screen "Rack 2" 640x480
   Button "Button_1" at 0,0 size 90x66; TextOff 'Rack 1'
      on Click: ActivateScreen("Rack 1", 0)
   Button "Button_2" at 130,0 size 90x66; TextOff 'Rack 2'
      on Click: ActivateScreen("Rack 2", 0)
   DateTimeField "Date/time field_1" at 444,15 size 177x31
   TextField "Text field_46" at 350,88 size 74x28; Text 'Rack 2'
   ScreenModuleView "RackSlot_1" at 562,360 size 44x36; Guid_{11997190-21654} '0'; ScreenModuleType ""
      on Guid_{11997190-21491}: function_efd93a16("RackSlotData", 0, 0, -1, -1, 1)
      Guid_{11997190-21133} <- "WarehouseData_Rack1{1}"
   ScreenModuleView "RackSlot_2" at 512,360 size 44x36; Guid_{11997190-21654} '0'; ScreenModuleType ""
      on Guid_{11997190-21491}: function_efd93a16("RackSlotData", 0, 0, -1, -1, 1)
      Guid_{11997190-21133} <- "WarehouseData_Rack1{1}"
   ScreenModuleView "RackSlot_3" at 562,360 size 44x36; Guid_{11997190-21654} '1'; Guid_{11997190-23841} '1'; ScreenModuleType ""
      on Guid_{11997190-21491}: SetTag("SelectedRack", 2); SetTag("SelectedSlot", 1); function_efd93a16("RackSlotData", 220, 150, -1, -1, 1)
      Guid_{11997190-21133} <- "WarehouseData_Rack2{1}"
   ScreenModuleView "RackSlot_4" at 512,360 size 44x36; Guid_{11997190-21654} '2'; Guid_{11997190-23841} '2'; ScreenModuleType ""
      on Guid_{11997190-21491}: SetTag("SelectedRack", 2); SetTag("SelectedSlot", 2); function_efd93a16("RackSlotData", 220, 150, -1, -1, 1)
      Guid_{11997190-21133} <- "WarehouseData_Rack2{2}"
   ScreenModuleView "RackSlot_5" at 462,360 size 44x36; Guid_{11997190-21654} '3'; Guid_{11997190-23841} '3'; ScreenModuleType ""
      on Guid_{11997190-21491}: SetTag("SelectedRack", 2); SetTag("SelectedSlot", 3); function_efd93a16("RackSlotData", 220, 150, -1, -1, 1)
      Guid_{11997190-21133} <- "WarehouseData_Rack2{3}"
   ScreenModuleView "RackSlot_6" at 412,360 size 44x36; Guid_{11997190-21654} '4'; Guid_{11997190-23841} '4'; ScreenModuleType ""
      on Guid_{11997190-21491}: SetTag("SelectedRack", 2); SetTag("SelectedSlot", 4); function_efd93a16("RackSlotData", 220, 150, -1, -1, 1)
      Guid_{11997190-21133} <- "WarehouseData_Rack2{4}"
   ScreenModuleView "RackSlot_7" at 362,360 size 44x36; Guid_{11997190-21654} '5'; Guid_{11997190-23841} '5'; ScreenModuleType ""
      on Guid_{11997190-21491}: SetTag("SelectedRack", 2); SetTag("SelectedSlot", 5); function_efd93a16("RackSlotData", 220, 150, -1, -1, 1)
      Guid_{11997190-21133} <- "WarehouseData_Rack2{5}"
   ScreenModuleView "RackSlot_8" at 312,360 size 44x36; Guid_{11997190-21654} '6'; Guid_{11997190-23841} '6'; ScreenModuleType ""
      on Guid_{11997190-21491}: SetTag("SelectedRack", 2); SetTag("SelectedSlot", 6); function_efd93a16("RackSlotData", 220, 150, -1, -1, 1)
      Guid_{11997190-21133} <- "WarehouseData_Rack2{6}"
   ScreenModuleView "RackSlot_9" at 262,360 size 44x36; Guid_{11997190-21654} '7'; Guid_{11997190-23841} '7'; ScreenModuleType ""
      on Guid_{11997190-21491}: SetTag("SelectedRack", 2); SetTag("SelectedSlot", 7); function_efd93a16("RackSlotData", 220, 150, -1, -1, 1)
      Guid_{11997190-21133} <- "WarehouseData_Rack2{7}"
   ScreenModuleView "RackSlot_10" at 212,360 size 44x36; Guid_{11997190-21654} '8'; Guid_{11997190-23841} '8'; ScreenModuleType ""
      on Guid_{11997190-21491}: SetTag("SelectedRack", 2); SetTag("SelectedSlot", 8); function_efd93a16("RackSlotData", 220, 150, -1, -1, 1)
      Guid_{11997190-21133} <- "WarehouseData_Rack2{8}"
   ScreenModuleView "RackSlot_11" at 162,360 size 44x36; Guid_{11997190-21654} '9'; Guid_{11997190-23841} '9'; ScreenModuleType ""
      on Guid_{11997190-21491}: SetTag("SelectedRack", 2); SetTag("SelectedSlot", 9); function_efd93a16("RackSlotData", 220, 150, -1, -1, 1)
      Guid_{11997190-21133} <- "WarehouseData_Rack2{9}"
   ScreenModuleView "RackSlot_12" at 562,315 size 44x36; Guid_{11997190-21654} '10'; Guid_{11997190-23841} '10'; ScreenModuleType ""
      on Guid_{11997190-21491}: SetTag("SelectedRack", 2); SetTag("SelectedSlot", 10); function_efd93a16("RackSlotData", 220, 150, -1, -1, 1)
      Guid_{11997190-21133} <- "WarehouseData_Rack2{10}"
   ScreenModuleView "RackSlot_13" at 512,315 size 44x36; Guid_{11997190-21654} '11'; Guid_{11997190-23841} '11'; ScreenModuleType ""
      on Guid_{11997190-21491}: SetTag("SelectedRack", 2); SetTag("SelectedSlot", 11); function_efd93a16("RackSlotData", 220, 150, -1, -1, 1)
      Guid_{11997190-21133} <- "WarehouseData_Rack2{11}"
   ScreenModuleView "RackSlot_14" at 462,315 size 44x36; Guid_{11997190-21654} '12'; Guid_{11997190-23841} '12'; ScreenModuleType ""
      on Guid_{11997190-21491}: SetTag("SelectedRack", 2); SetTag("SelectedSlot", 12); function_efd93a16("RackSlotData", 220, 150, -1, -1, 1)
      Guid_{11997190-21133} <- "WarehouseData_Rack2{12}"
   ScreenModuleView "RackSlot_15" at 412,315 size 44x36; Guid_{11997190-21654} '13'; Guid_{11997190-23841} '13'; ScreenModuleType ""
      on Guid_{11997190-21491}: SetTag("SelectedRack", 2); SetTag("SelectedSlot", 13); function_efd93a16("RackSlotData", 220, 150, -1, -1, 1)
      Guid_{11997190-21133} <- "WarehouseData_Rack2{13}"
   ScreenModuleView "RackSlot_16" at 362,315 size 44x36; Guid_{11997190-21654} '14'; Guid_{11997190-23841} '14'; ScreenModuleType ""
      on Guid_{11997190-21491}: SetTag("SelectedRack", 2); SetTag("SelectedSlot", 14); function_efd93a16("RackSlotData", 220, 150, -1, -1, 1)
      Guid_{11997190-21133} <- "WarehouseData_Rack2{14}"
   ScreenModuleView "RackSlot_17" at 312,315 size 44x36; Guid_{11997190-21654} '15'; Guid_{11997190-23841} '15'; ScreenModuleType ""
      on Guid_{11997190-21491}: SetTag("SelectedRack", 2); SetTag("SelectedSlot", 15); function_efd93a16("RackSlotData", 220, 150, -1, -1, 1)
      Guid_{11997190-21133} <- "WarehouseData_Rack2{15}"
   ScreenModuleView "RackSlot_18" at 262,315 size 44x36; Guid_{11997190-21654} '16'; Guid_{11997190-23841} '16'; ScreenModuleType ""
      on Guid_{11997190-21491}: SetTag("SelectedRack", 2); SetTag("SelectedSlot", 16); function_efd93a16("RackSlotData", 220, 150, -1, -1, 1)
      Guid_{11997190-21133} <- "WarehouseData_Rack2{16}"
   ScreenModuleView "RackSlot_19" at 212,315 size 44x36; Guid_{11997190-21654} '17'; Guid_{11997190-23841} '17'; ScreenModuleType ""
      on Guid_{11997190-21491}: SetTag("SelectedRack", 2); SetTag("SelectedSlot", 17); function_efd93a16("RackSlotData", 220, 150, -1, -1, 1)
      Guid_{11997190-21133} <- "WarehouseData_Rack2{17}"
   ScreenModuleView "RackSlot_20" at 162,315 size 44x36; Guid_{11997190-21654} '18'; Guid_{11997190-23841} '18'; ScreenModuleType ""
      on Guid_{11997190-21491}: SetTag("SelectedRack", 2); SetTag("SelectedSlot", 18); function_efd93a16("RackSlotData", 220, 150, -1, -1, 1)
      Guid_{11997190-21133} <- "WarehouseData_Rack2{18}"
   ScreenModuleView "RackSlot_21" at 562,270 size 44x36; Guid_{11997190-21654} '19'; Guid_{11997190-23841} '19'; ScreenModuleType ""
      on Guid_{11997190-21491}: SetTag("SelectedRack", 2); SetTag("SelectedSlot", 19); function_efd93a16("RackSlotData", 220, 150, -1, -1, 1)
      Guid_{11997190-21133} <- "WarehouseData_Rack2{19}"
   ScreenModuleView "RackSlot_22" at 512,270 size 44x36; Guid_{11997190-21654} '20'; Guid_{11997190-23841} '20'; ScreenModuleType ""
      on Guid_{11997190-21491}: SetTag("SelectedRack", 2); SetTag("SelectedSlot", 20); function_efd93a16("RackSlotData", 220, 150, -1, -1, 1)
      Guid_{11997190-21133} <- "WarehouseData_Rack2{20}"
   ScreenModuleView "RackSlot_23" at 462,270 size 44x36; Guid_{11997190-21654} '21'; Guid_{11997190-23841} '21'; ScreenModuleType ""
      on Guid_{11997190-21491}: SetTag("SelectedRack", 2); SetTag("SelectedSlot", 21); function_efd93a16("RackSlotData", 220, 150, -1, -1, 1)
      Guid_{11997190-21133} <- "WarehouseData_Rack2{21}"
   ScreenModuleView "RackSlot_24" at 412,270 size 44x36; Guid_{11997190-21654} '22'; Guid_{11997190-23841} '22'; ScreenModuleType ""
      on Guid_{11997190-21491}: SetTag("SelectedRack", 2); SetTag("SelectedSlot", 22); function_efd93a16("RackSlotData", 220, 150, -1, -1, 1)
      Guid_{11997190-21133} <- "WarehouseData_Rack2{22}"
   ScreenModuleView "RackSlot_25" at 362,270 size 44x36; Guid_{11997190-21654} '23'; Guid_{11997190-23841} '23'; ScreenModuleType ""
      on Guid_{11997190-21491}: SetTag("SelectedRack", 2); SetTag("SelectedSlot", 23); function_efd93a16("RackSlotData", 220, 150, -1, -1, 1)
      Guid_{11997190-21133} <- "WarehouseData_Rack2{23}"
   ScreenModuleView "RackSlot_26" at 312,270 size 44x36; Guid_{11997190-21654} '24'; Guid_{11997190-23841} '24'; ScreenModuleType ""
      on Guid_{11997190-21491}: SetTag("SelectedRack", 2); SetTag("SelectedSlot", 24); function_efd93a16("RackSlotData", 220, 150, -1, -1, 1)
      Guid_{11997190-21133} <- "WarehouseData_Rack2{24}"
   ScreenModuleView "RackSlot_27" at 262,270 size 44x36; Guid_{11997190-21654} '25'; Guid_{11997190-23841} '25'; ScreenModuleType ""
      on Guid_{11997190-21491}: SetTag("SelectedRack", 2); SetTag("SelectedSlot", 25); function_efd93a16("RackSlotData", 220, 150, -1, -1, 1)
      Guid_{11997190-21133} <- "WarehouseData_Rack2{25}"
   ScreenModuleView "RackSlot_28" at 212,270 size 44x36; Guid_{11997190-21654} '26'; Guid_{11997190-23841} '26'; ScreenModuleType ""
      on Guid_{11997190-21491}: SetTag("SelectedRack", 2); SetTag("SelectedSlot", 26); function_efd93a16("RackSlotData", 220, 150, -1, -1, 1)
      Guid_{11997190-21133} <- "WarehouseData_Rack2{26}"
   ScreenModuleView "RackSlot_29" at 162,270 size 44x36; Guid_{11997190-21654} '27'; Guid_{11997190-23841} '27'; ScreenModuleType ""
      on Guid_{11997190-21491}: SetTag("SelectedRack", 2); SetTag("SelectedSlot", 27); function_efd93a16("RackSlotData", 220, 150, -1, -1, 1)
      Guid_{11997190-21133} <- "WarehouseData_Rack2{27}"
   ScreenModuleView "RackSlot_30" at 562,225 size 44x36; Guid_{11997190-21654} '28'; Guid_{11997190-23841} '28'; ScreenModuleType ""
      on Guid_{11997190-21491}: SetTag("SelectedRack", 2); SetTag("SelectedSlot", 28); function_efd93a16("RackSlotData", 220, 150, -1, -1, 1)
      Guid_{11997190-21133} <- "WarehouseData_Rack2{28}"
   ScreenModuleView "RackSlot_31" at 512,225 size 44x36; Guid_{11997190-21654} '29'; Guid_{11997190-23841} '29'; ScreenModuleType ""
      on Guid_{11997190-21491}: SetTag("SelectedRack", 2); SetTag("SelectedSlot", 29); function_efd93a16("RackSlotData", 220, 150, -1, -1, 1)
      Guid_{11997190-21133} <- "WarehouseData_Rack2{29}"
   ScreenModuleView "RackSlot_32" at 462,225 size 44x36; Guid_{11997190-21654} '30'; Guid_{11997190-23841} '30'; ScreenModuleType ""
      on Guid_{11997190-21491}: SetTag("SelectedRack", 2); SetTag("SelectedSlot", 30); function_efd93a16("RackSlotData", 220, 150, -1, -1, 1)
      Guid_{11997190-21133} <- "WarehouseData_Rack2{30}"
   ScreenModuleView "RackSlot_33" at 412,225 size 44x36; Guid_{11997190-21654} '31'; Guid_{11997190-23841} '31'; ScreenModuleType ""
      on Guid_{11997190-21491}: SetTag("SelectedRack", 2); SetTag("SelectedSlot", 31); function_efd93a16("RackSlotData", 220, 150, -1, -1, 1)
      Guid_{11997190-21133} <- "WarehouseData_Rack2{31}"
   ScreenModuleView "RackSlot_34" at 362,225 size 44x36; Guid_{11997190-21654} '32'; Guid_{11997190-23841} '32'; ScreenModuleType ""
      on Guid_{11997190-21491}: SetTag("SelectedRack", 2); SetTag("SelectedSlot", 32); function_efd93a16("RackSlotData", 220, 150, -1, -1, 1)
      Guid_{11997190-21133} <- "WarehouseData_Rack2{32}"
   ScreenModuleView "RackSlot_35" at 312,225 size 44x36; Guid_{11997190-21654} '33'; Guid_{11997190-23841} '33'; ScreenModuleType ""
      on Guid_{11997190-21491}: SetTag("SelectedRack", 2); SetTag("SelectedSlot", 33); function_efd93a16("RackSlotData", 220, 150, -1, -1, 1)
      Guid_{11997190-21133} <- "WarehouseData_Rack2{33}"
   ScreenModuleView "RackSlot_36" at 262,225 size 44x36; Guid_{11997190-21654} '34'; Guid_{11997190-23841} '34'; ScreenModuleType ""
      on Guid_{11997190-21491}: SetTag("SelectedRack", 2); SetTag("SelectedSlot", 34); function_efd93a16("RackSlotData", 220, 150, -1, -1, 1)
      Guid_{11997190-21133} <- "WarehouseData_Rack2{34}"
   ScreenModuleView "RackSlot_37" at 212,225 size 44x36; Guid_{11997190-21654} '35'; Guid_{11997190-23841} '35'; ScreenModuleType ""
      on Guid_{11997190-21491}: SetTag("SelectedRack", 2); SetTag("SelectedSlot", 36); function_efd93a16("RackSlotData", 220, 150, -1, -1, 1)
      Guid_{11997190-21133} <- "WarehouseData_Rack2{35}"
   ScreenModuleView "RackSlot_38" at 162,225 size 44x36; Guid_{11997190-21654} '36'; Guid_{11997190-23841} '36'; ScreenModuleType ""
      on Guid_{11997190-21491}: SetTag("SelectedRack", 2); SetTag("SelectedSlot", 36); function_efd93a16("RackSlotData", 220, 150, -1, -1, 1)
      Guid_{11997190-21133} <- "WarehouseData_Rack2{36}"
   ScreenModuleView "RackSlot_39" at 562,180 size 44x36; Guid_{11997190-21654} '37'; Guid_{11997190-23841} '37'; ScreenModuleType ""
      on Guid_{11997190-21491}: SetTag("SelectedRack", 2); SetTag("SelectedSlot", 37); function_efd93a16("RackSlotData", 220, 150, -1, -1, 1)
      Guid_{11997190-21133} <- "WarehouseData_Rack2{37}"
   ScreenModuleView "RackSlot_40" at 512,180 size 44x36; Guid_{11997190-21654} '38'; Guid_{11997190-23841} '38'; ScreenModuleType ""
      on Guid_{11997190-21491}: SetTag("SelectedRack", 2); SetTag("SelectedSlot", 38); function_efd93a16("RackSlotData", 220, 150, -1, -1, 1)
      Guid_{11997190-21133} <- "WarehouseData_Rack2{38}"
   ScreenModuleView "RackSlot_41" at 462,180 size 44x36; Guid_{11997190-21654} '39'; Guid_{11997190-23841} '39'; ScreenModuleType ""
      on Guid_{11997190-21491}: SetTag("SelectedRack", 2); SetTag("SelectedSlot", 39); function_efd93a16("RackSlotData", 220, 150, -1, -1, 1)
      Guid_{11997190-21133} <- "WarehouseData_Rack2{39}"
   ScreenModuleView "RackSlot_42" at 412,180 size 44x36; Guid_{11997190-21654} '40'; Guid_{11997190-23841} '40'; ScreenModuleType ""
      on Guid_{11997190-21491}: SetTag("SelectedRack", 2); SetTag("SelectedSlot", 40); function_efd93a16("RackSlotData", 220, 150, -1, -1, 1)
      Guid_{11997190-21133} <- "WarehouseData_Rack2{40}"
   ScreenModuleView "RackSlot_43" at 362,180 size 44x36; Guid_{11997190-21654} '41'; Guid_{11997190-23841} '41'; ScreenModuleType ""
      on Guid_{11997190-21491}: SetTag("SelectedRack", 2); SetTag("SelectedSlot", 41); function_efd93a16("RackSlotData", 220, 150, -1, -1, 1)
      Guid_{11997190-21133} <- "WarehouseData_Rack2{41}"
   ScreenModuleView "RackSlot_44" at 312,180 size 44x36; Guid_{11997190-21654} '42'; Guid_{11997190-23841} '42'; ScreenModuleType ""
      on Guid_{11997190-21491}: SetTag("SelectedRack", 2); SetTag("SelectedSlot", 42); function_efd93a16("RackSlotData", 220, 150, -1, -1, 1)
      Guid_{11997190-21133} <- "WarehouseData_Rack2{42}"
   ScreenModuleView "RackSlot_45" at 262,180 size 44x36; Guid_{11997190-21654} '43'; Guid_{11997190-23841} '43'; ScreenModuleType ""
      on Guid_{11997190-21491}: SetTag("SelectedRack", 2); SetTag("SelectedSlot", 43); function_efd93a16("RackSlotData", 220, 150, -1, -1, 1)
      Guid_{11997190-21133} <- "WarehouseData_Rack2{43}"
   ScreenModuleView "RackSlot_46" at 212,180 size 44x36; Guid_{11997190-21654} '44'; Guid_{11997190-23841} '44'; ScreenModuleType ""
      on Guid_{11997190-21491}: SetTag("SelectedRack", 2); SetTag("SelectedSlot", 44); function_efd93a16("RackSlotData", 220, 150, -1, -1, 1)
      Guid_{11997190-21133} <- "WarehouseData_Rack2{44}"
   ScreenModuleView "RackSlot_47" at 162,180 size 44x36; Guid_{11997190-21654} '45'; Guid_{11997190-23841} '45'; ScreenModuleType ""
      on Guid_{11997190-21491}: SetTag("SelectedRack", 2); SetTag("SelectedSlot", 45); function_efd93a16("RackSlotData", 220, 150, -1, -1, 1)
      Guid_{11997190-21133} <- "WarehouseData_Rack2{45}"
   ScreenModuleView "RackSlot_48" at 562,135 size 44x36; Guid_{11997190-21654} '46'; Guid_{11997190-23841} '46'; ScreenModuleType ""
      on Guid_{11997190-21491}: SetTag("SelectedRack", 2); SetTag("SelectedSlot", 46); function_efd93a16("RackSlotData", 220, 150, -1, -1, 1)
      Guid_{11997190-21133} <- "WarehouseData_Rack2{46}"
   ScreenModuleView "RackSlot_49" at 512,135 size 44x36; Guid_{11997190-21654} '47'; Guid_{11997190-23841} '47'; ScreenModuleType ""
      on Guid_{11997190-21491}: SetTag("SelectedRack", 2); SetTag("SelectedSlot", 47); function_efd93a16("RackSlotData", 220, 150, -1, -1, 1)
      Guid_{11997190-21133} <- "WarehouseData_Rack2{47}"
   ScreenModuleView "RackSlot_50" at 462,135 size 44x36; Guid_{11997190-21654} '48'; Guid_{11997190-23841} '48'; ScreenModuleType ""
      on Guid_{11997190-21491}: SetTag("SelectedRack", 2); SetTag("SelectedSlot", 48); function_efd93a16("RackSlotData", 220, 150, -1, -1, 1)
      Guid_{11997190-21133} <- "WarehouseData_Rack2{48}"
   ScreenModuleView "RackSlot_51" at 412,135 size 44x36; Guid_{11997190-21654} '49'; Guid_{11997190-23841} '49'; ScreenModuleType ""
      on Guid_{11997190-21491}: SetTag("SelectedRack", 2); SetTag("SelectedSlot", 49); function_efd93a16("RackSlotData", 220, 150, -1, -1, 1)
      Guid_{11997190-21133} <- "WarehouseData_Rack2{49}"
   ScreenModuleView "RackSlot_52" at 362,135 size 44x36; Guid_{11997190-21654} '50'; Guid_{11997190-23841} '50'; ScreenModuleType ""
      on Guid_{11997190-21491}: SetTag("SelectedRack", 2); SetTag("SelectedSlot", 50); function_efd93a16("RackSlotData", 220, 150, -1, -1, 1)
      Guid_{11997190-21133} <- "WarehouseData_Rack2{50}"
   ScreenModuleView "RackSlot_53" at 312,135 size 44x36; Guid_{11997190-21654} '51'; Guid_{11997190-23841} '51'; ScreenModuleType ""
      on Guid_{11997190-21491}: SetTag("SelectedRack", 2); SetTag("SelectedSlot", 51); function_efd93a16("RackSlotData", 220, 150, -1, -1, 1)
      Guid_{11997190-21133} <- "WarehouseData_Rack2{51}"
   ScreenModuleView "RackSlot_54" at 262,135 size 44x36; Guid_{11997190-21654} '52'; Guid_{11997190-23841} '52'; ScreenModuleType ""
      on Guid_{11997190-21491}: SetTag("SelectedRack", 2); SetTag("SelectedSlot", 52); function_efd93a16("RackSlotData", 220, 150, -1, -1, 1)
      Guid_{11997190-21133} <- "WarehouseData_Rack2{52}"
   ScreenModuleView "RackSlot_55" at 212,135 size 44x36; Guid_{11997190-21654} '53'; Guid_{11997190-23841} '53'; ScreenModuleType ""
      on Guid_{11997190-21491}: SetTag("SelectedRack", 2); SetTag("SelectedSlot", 53); function_efd93a16("RackSlotData", 220, 150, -1, -1, 1)
      Guid_{11997190-21133} <- "WarehouseData_Rack2{53}"
   ScreenModuleView "RackSlot_56" at 162,135 size 44x36; Guid_{11997190-21654} '54'; Guid_{11997190-23841} '54'; ScreenModuleType ""
      on Guid_{11997190-21491}: SetTag("SelectedRack", 2); SetTag("SelectedSlot", 54); function_efd93a16("RackSlotData", 220, 150, -1, -1, 1)
      Guid_{11997190-21133} <- "WarehouseData_Rack2{54}"
   TextField "Text field_1" at 17,171 size 106x22; Text 'Crane Status:'
   TextField "Text field_2" at 17,360 size 113x22; Text 'Both racks full'
      Visibility <- "RacksFull"
   TextField "Text field_4" at 15,121 size 15x22; Text 'Text'
   TextField "Text field_3" at 17,193 size 70x18; Text 'Text'
   TextField "Text field_5" at 17,261 size 119x22; Text 'Occupied slots:'
   TextField "Text field_6" at 36,283 size 28x18; Text '/ 54'
   TextField "Text field_7" at 17,283 size 29x18; Text 'Text'
   Button "Button_3" at 17,104 size 54x39; TextOff 'START'
      on Press: SetBit("StartCmd")
      on Release: ResetBit("StartCmd")
   Button "Button_4" at 80,104 size 54x39; TextOff 'STOP'
      on Press: SetBit("StopCmd")
      on Release: ResetBit("StopCmd")

VB script "VBFunction_1"
   'Tip:
   ' 1. Use the <CTRL+SPACE> or <CTRL+I> shortcut to open a list of all objects and functions
   ' 2. Write the code using the HMI Runtime object.
   '  Example: HmiRuntime.Screens("Screen_1").
   ' 3. Use the <CTRL+J> shortcut to create an object reference.
   'Write the code as of this position:
*)

(* ===== HMI "HMI_RT_1" =====

ScreenModuleEditorView "RackSlot" 640x480
   Rectangle "Rectangle_1" at 348,118 size 50x40
      Appearance <- "WarehouseSlots.Status"
   TextField "Text field_1" at 363,127 size 15x22; Text '0'
   Button "Button_1" at 348,118 size 50x40; TextOff 's'
*)